(*
.. admonition:: And, by the way...

   You can make up your own admonition too.
*)

FUNCTION_BLOCK FB_Libdoc_GenericNotes
VAR_INPUT
    nVarA : INT;
    nVarB : INT;
END_VAR
VAR_OUTPUT
    nSum : INT;
END_VAR
VAR
END_VAR

END_FUNCTION_BLOCK

(* stored: Version 1.1.0.1, ProductVersion 3.1.4022.18
   POU FB_Libdoc_GenericNotes: Id {d6ae01ea-f028-4cf4-9848-81962ce46acb}, SpecialFunc None *)
